(* IEC 61131-3 sources: llm-plc-st-eval/data/processed_definitivo/claude-sonnet-4-6/C7/zero_shot, 3 files *)

(* ---- ejec_1.st ---- *)
FUNCTION_BLOCK FB_Contador
VAR_INPUT
    sensorPieza : BOOL; (* Sensor de detección de pieza *)
    btnReset    : BOOL; (* Botón de reset del contador *)
END_VAR

VAR_OUTPUT
    loteListo : BOOL; (* Indica que el lote de 12 piezas está completo *)
    cuenta    : INT;  (* Valor actual del contador *)
END_VAR

VAR
    C1 : CTU; (* Contador ascendente IEC 61131-3 *)
END_VAR

(* -------------------------------------------------------
   Rama 1: Contador ascendente C1
   CU  <- sensorPieza (flanco ascendente cuenta una pieza)
   RESET <- btnReset  (reinicia el contador)
   PV  = 12           (tamaño del lote)
------------------------------------------------------- *)
C1(
    CU    := sensorPieza,
    RESET := btnReset,
    PV    := 12
);

(* -------------------------------------------------------
   Rama 2: Activar loteListo cuando el contador alcanza PV
   Equivale al contacto normalmente abierto de C1.Q
   alimentando la bobina loteListo
------------------------------------------------------- *)
loteListo := C1.Q;

(* -------------------------------------------------------
   Rama 3: Transferir el valor actual del contador
   a la variable de salida cuenta
------------------------------------------------------- *)
cuenta := C1.CV;

END_FUNCTION_BLOCK

(* ---- ejec_2.st ---- *)
FUNCTION_BLOCK FB_Contador
VAR_INPUT
    sensorPieza : BOOL; (* Sensor de detección de pieza *)
    btnReset    : BOOL; (* Botón de reset del contador *)
END_VAR

VAR_OUTPUT
    loteListo : BOOL; (* Indica que el lote de 12 piezas está completo *)
    cuenta    : INT;  (* Valor actual del contador *)
END_VAR

VAR
    C1 : CTU; (* Contador ascendente IEC 61131-3 *)
END_VAR

(* -------------------------------------------------------
   Rama 1: Contador ascendente C1
   CU  <- sensorPieza (flanco ascendente cuenta una pieza)
   R   <- btnReset    (reset del contador)
   PV  = 12          (valor preestablecido del lote)
   ------------------------------------------------------- *)
C1(
    CU := sensorPieza,
    R  := btnReset,
    PV := 12
);

(* -------------------------------------------------------
   Rama 2: Bobina loteListo
   Se activa cuando C1.Q = TRUE (CV >= PV)
   ------------------------------------------------------- *)
loteListo := C1.Q;

(* -------------------------------------------------------
   Rama 3: Transferencia del valor actual a cuenta
   ------------------------------------------------------- *)
cuenta := C1.CV;
END_FUNCTION_BLOCK

(* ---- ejec_3.st ---- *)
FUNCTION_BLOCK FB_Contador
VAR_INPUT
    sensorPieza : BOOL; (* Sensor de detección de pieza (contacto NA) *)
    btnReset    : BOOL; (* Botón de reset del contador (contacto NA) *)
END_VAR

VAR_OUTPUT
    loteListo : BOOL; (* Activa cuando se completa el lote (C1.Q) *)
    cuenta    : INT;  (* Valor actual del contador (C1.CV) *)
END_VAR

VAR
    C1 : CTU; (* Contador ascendente IEC 61131-3 *)
END_VAR

(* ---------------------------------------------------------------
   Rama 1: sensorPieza -> CU de C1 | btnReset -> RESET de C1
   Rama 2: C1.Q -> loteListo
   Rama 3: C1.CV -> cuenta
--------------------------------------------------------------- *)

(* Rama 1: llamada al contador CTU *)
C1(
    CU    := sensorPieza, (* Flanco ascendente de sensorPieza incrementa el contador *)
    RESET := btnReset,    (* btnReset pone CV a 0 y Q a FALSE *)
    PV    := 12           (* Valor preestablecido del lote *)
);

(* Rama 2: la salida Q del contador activa loteListo *)
loteListo := C1.Q;

(* Rama 3: transferencia del valor actual a la variable cuenta *)
cuenta := C1.CV;
